Fanuc KAREL source: kb00161.KL

-- PROVISIONAL review KL for V770-1; original PC SHA256 b22cc1e3fc4768af5cc0d6cf06efe6dab95c196adad1a4bf655397b2d720d209
-- Incomplete behavior may be omitted. Consult companion uncertainty JSON. Do not deploy.
PROGRAM KB00161
%NOLOCKGROUP
BEGIN
  -- UNRESOLVED_PC offsets 5-12; opcodes 9D,23
  -- UNRESOLVED_PC offsets 17-24; opcodes 9D,23
  -- UNRESOLVED_PC offsets 29-59; opcodes 27,22,22,1C,22,27,9D,31
  -- UNRESOLVED_PC offsets 64-68; opcodes 7F
END KB00161
